{attribute 'linkalways'}
{attribute 'no_explicit_call' := 'This FB is a CLASS and must be accessed using methods or properties'}
{attribute 'enable_dynamic_creation'}
FUNCTION_BLOCK Node_F_VN_CopyIntoDisplayableImageExp EXTENDS VisionNode
VAR
    ipSrcImage : _ITcVnImage;
    ipDestImage : _ITcVnDisplayableImage;
    nTimestamp : _LINT(0);
    hrPrev : _HRESULT(S_OK);
    hresult : _HRESULT(S_OK);
END_VAR

METHOD PUBLIC Clone : I_Node
VAR
    pNode : POINTER TO Node_F_VN_CopyIntoDisplayableImageExp;
END_VAR
pNode := __NEW(Node_F_VN_CopyIntoDisplayableImageExp);
Clone := pNode^;
END_METHOD

METHOD FB_init : BOOL
VAR_INPUT
    bInitRetains : BOOL;
    bInCopyCode : BOOL;
END_VAR
AddInput('ipSrcImage', ipSrcImage);
AddParameter('nTimestamp', nTimestamp);
AddInput('hrPrev', hrPrev);
AddOutput('ipDestImage', ipDestImage);
AddOutput('hresult', hresult);
END_METHOD

METHOD PROTECTED OnExecute
hresult.Value := F_VN_CopyIntoDisplayableImageExp(
    ipSrcImage := ipSrcImage.Value,
    ipDestImage := ipDestImage.Value,
    nTimestamp := nTimestamp.Value,
    hrPrev := hrPrev.Value);
END_METHOD

METHOD PUBLIC PreExecutionCheck
VAR_INPUT
    Check : I_PreExecutionChecks;
END_VAR
Check.IsTrue(ipSrcImage.IsValid, 'ipSrcImage must contain an image');
END_METHOD

END_FUNCTION_BLOCK

(* stored: Version 1.1.0.1, ProductVersion 3.1.4026.19
   POU Node_F_VN_CopyIntoDisplayableImageExp: Id {f6d1a4a8-83b1-4ce3-9636-921a7fa74d26}, SpecialFunc None
   Folder Constructor: Id {96ca97ff-9096-4d73-ad6f-45c90b1feaf8}
   Method Clone: Id {7598b5bf-66e5-4262-81bd-3c0d7d65ae43}
   Method FB_init: Id {8a066b0e-dd8a-45af-aba9-b9abead7dc39}
   Method OnExecute: Id {d99ccda3-c8ad-4675-8b54-69d5100ca439}
   Method PreExecutionCheck: Id {1ae8ac68-171e-46bd-b4ba-1b108720329a} *)
